FUNCTION_BLOCK FB_CellDevices
VAR
    FeedAxis : FB_SimAxis;
    TrackMover : FB_SimAxis;
    ShuttleX : FB_SimAxis;
    ShuttleY : FB_SimAxis;
    Camera : FB_SealInspection;
END_VAR
VAR_OUTPUT
    Indexing : BOOL;
    Rejected : DINT;
END_VAR
VAR_INPUT
    MissingSeal : BOOL;
END_VAR

METHOD ResetDevices
FeedAxis.Home();
TrackMover.Home();
ShuttleX.Home();
ShuttleY.Home();
Camera.ClearResult();
Indexing := FALSE;
END_METHOD

METHOD ProcessStation
VAR_INPUT
    Station : DINT;
    Phase : DINT;
END_VAR
CASE Station OF
    1: // Servo meters a 180 mm blank.
        FeedAxis.MoveToward(180, 2);
    4: // Trigger once when the closing platen reaches its forward limit.
        IF Phase >= 100 THEN Camera.Inspect(MissingSeal); END_IF
    5: // Route the sealed carton to one of two discharge lanes.
        ShuttleX.MoveToward(240, 2);
        ShuttleY.MoveToward(SEL(Camera.Verdict = 1, -120, 120), 2);
END_CASE
END_METHOD

METHOD IndexToNext : BOOL
VAR_INPUT
    Station : DINT;
END_VAR
IndexToNext := TrackMover.MoveToward(Station * 560, 8);
Indexing := NOT IndexToNext;
END_METHOD

METHOD ReadyToLeave : BOOL
VAR_INPUT
    Station : DINT;
END_VAR
CASE Station OF
    1: ReadyToLeave := FeedAxis.PositionMm = 180;
    4: ReadyToLeave := Camera.Verdict <> 0;
    5: ReadyToLeave := (ShuttleX.PositionMm = 240) AND
           (ShuttleY.PositionMm = SEL(Camera.Verdict = 1, -120, 120));
ELSE
    ReadyToLeave := TRUE;
END_CASE
END_METHOD

METHOD FinishCarton : BOOL
FinishCarton := Camera.Verdict = 1;
IF NOT FinishCarton THEN Rejected := Rejected + 1; END_IF
END_METHOD

METHOD Publish
VAR_IN_OUT
    Words : ARRAY[0..105] OF DINT;
END_VAR
Words[11] := FeedAxis.PositionMm;
Words[12] := TrackMover.PositionMm;
Words[13] := ShuttleX.PositionMm;
Words[14] := ShuttleY.PositionMm;
Words[15] := Camera.Verdict;
Words[16] := Rejected;
Words[17] := BOOL_TO_DINT(MissingSeal);
Words[18] := BOOL_TO_DINT(Indexing);
Words[19] := Camera.BrightSamples;
END_METHOD

END_FUNCTION_BLOCK

(* stored: Version 1.1.0.1
   POU FB_CellDevices: Id {69468DC3-8A7A-45D7-9465-000000000007}
   Method ResetDevices: Id {69468DC3-8A7A-45D7-9465-000000000008}
   Method ProcessStation: Id {69468DC3-8A7A-45D7-9465-000000000009}
   Method IndexToNext: Id {69468DC3-8A7A-45D7-9465-000000000010}
   Method ReadyToLeave: Id {0DFB410B-908E-4365-B964-B1C23F60891C}
   Method FinishCarton: Id {69468DC3-8A7A-45D7-9465-000000000011}
   Method Publish: Id {69468DC3-8A7A-45D7-9465-000000000012} *)
